(* PLC project , CODESYS CODESYS V3.5 SP16 Patch 4 *)
(* stored: creationDateTime 2022-07-19T13:27:04.6322144, modificationDateTime 2021-08-16T16:25:27.2929866 *)

FUNCTION_BLOCK ccsSafeCraneNumberSuperv
  VAR_INPUT
    in_CraneNoSet1 : WORD;  (* First crane number *)
    in_CraneNoSet2 : WORD;  (* Second crane number *)
  END_VAR
  VAR_OUTPUT
    out_S_CraneNoSupervOk : BOOL;  (* Crane numbers match and are not an empty word *)
    out_S_CraneNo : WORD;  (* A safe crane number. If crane numbers missmatch, this word is set to an empty word *)
  END_VAR
  VAR
    EmptyWord : WORD;
  END_VAR

            out_S_CraneNoSupervOk :=
	(in_CraneNoSet1 = in_CraneNoSet2)
	AND (in_CraneNoSet1 <> EmptyWord);

IF out_S_CraneNoSupervOk THEN
	out_S_CraneNo := in_CraneNoSet1;
ELSE
	out_S_CraneNo := EmptyWord;
END_IF
          
END_FUNCTION_BLOCK
